// TwinCAT 3 PLC project CMoLib
// ProgramVersion: 3.1.4024.0
// libraries:
//   Tc2_Standard, * (Beckhoff Automation GmbH)
//   Tc2_System, * (Beckhoff Automation GmbH)
//   Tc2_Utilities, * (Beckhoff Automation GmbH)
//   Tc3_Module, * (Beckhoff Automation GmbH)
// project tree:
//   DUTs/ CMoDateTime.TcDUT, CMoDateTimeString.TcDUT, CMoFramework.TcDUT, CMoHalDigitalInput.TcDUT, CMoHalDigitalOutput.TcDUT, CMoInterlock.TcDUT
//   GVLs/ GVL.TcGVL
//   / PlcTask.TcTTO
//   POUs/ CMoDateTimeToString.TcPOU, CMoDiffTime.TcPOU, CMoDigitalInput.TcPOU, CMoDigitalOutput.TcPOU, CMoElapsedTime.TcPOU, CMoEvalInterlock.TcPOU, CMoGetLocalDateTime.TcPOU, CMoGetUTCDateTime.TcPOU, CMoMainRuntime.TcPOU, CMoRandom.TcPOU, MAIN.TcPOU
// real-time tasks:
//   TASK PlcTask: cycle T#5ms, priority 20, ADS port 350

CONFIGURATION CMoLib
    RESOURCE PLC ON TwinCAT3
        TASK PlcTask(INTERVAL := T#5ms, PRIORITY := 20);
        PROGRAM MAIN WITH PlcTask : MAIN;
    END_RESOURCE
END_CONFIGURATION

// ---- DUTs/CMoDateTime.TcDUT
// CMoDateTime — Date and Time Structure
// CMo Library v1.0 — Cristian Mori
// TwinCAT / IEC 61131-3 Structured Text

TYPE CMoDateTime :
STRUCT
    RawDateTime     : ARRAY[0..6] OF DINT;  // Platform-native wall clock data
    Year            : DINT;
    Month           : DINT;     // 1-12
    Day             : DINT;     // 1-31
    Hour            : DINT;     // 0-23
    Minute          : DINT;     // 0-59
    Second          : DINT;     // 0-59
    MicroSecond     : DINT;     // 0-999999
    IsLocal         : BOOL;     // TRUE = local time, FALSE = UTC
END_STRUCT
END_TYPE

// ---- DUTs/CMoDateTimeString.TcDUT
// CMoDateTimeString — HMI-Readable Date/Time Strings
// CMo Library v1.0 — Cristian Mori

TYPE CMoDateTimeString :
STRUCT
    TimeString      : STRING(16);   // "HH:MM:SS"
    DateString      : STRING(16);   // "YYYY-MM-DD"
    HMIString       : STRING(32);   // "YYYY-MM-DD HH:MM:SS"
END_STRUCT
END_TYPE

// ---- DUTs/CMoFramework.TcDUT
// CMoCommon — Shared System Context
// CMo Library v1.0 — Cristian Mori
//
// One instance per PLC. Passed as VAR_IN_OUT to every FB.
// Temp* fields are scratch accumulators: reset each scan by CMoMasterTask,
// set by individual FBs, then latched into final fields next scan.

TYPE CMoFramework :
STRUCT
    // ---- Alarm rollup flags ----
    AnyAudibleOn            : BOOL;
    AnyAudibleOnLastScan        : BOOL;
    AnyAlarmActive          : BOOL;
    AnyAlarmActiveLastScan      : BOOL;
    AnyWarningActive        : BOOL;
    AnyWarningActiveLastScan    : BOOL;
    AnyFaultActive          : BOOL;
    AnyFaultActiveLastScan      : BOOL;
    AnyCriticalActive       : BOOL;
    AnyCriticalActiveLastScan   : BOOL;

    // ---- Simulation / Hand detection ----
    AnySimulationOn         : BOOL;
    AnySimulationOnLastScan     : BOOL;
    AnyHandOn               : BOOL;
    AnyHandOnLastScan           : BOOL;

    // ---- HMI commands ----
    SilenceCmd              : BOOL;     // HMI silence button (momentary)
    GlobalAlmRstCmd         : BOOL;     // HMI global alarm reset (momentary)
    GlobalAlmRstEn          : BOOL;     // Enable global alarm reset

    // ---- System modes ----
    SimulationEnabled       : BOOL;     // Master simulation enable
    EmulationEnabled        : BOOL;     // Running on emulated controller
    MaintenanceEnabled      : BOOL;     // Enables Hand mode

    // ---- Tick timers (pulse TRUE for one scan) ----
    Tick100ms               : BOOL;
    Tick1s                  : BOOL;
    Tick10s                 : BOOL;

    // ---- Blinker signals (toggle on/off) ----
	Blink100ms				: BOOL;
    Blink250ms              : BOOL;
    Blink500ms              : BOOL;
    Blink1s                 : BOOL;
    Blink2s                 : BOOL;

    // ---- System flags ----
    InhibitAlarms           : BOOL;     // Corporate alarm inhibit
    AlwaysTrue              : BOOL;     // Constant TRUE
    AlwaysFalse             : BOOL;     // Constant FALSE
  

    // ---- Counters ----
    ApplicationCount        : DINT;
    AlarmCount              : INT;
    TempAlarmCount          : INT;
    FreeRunningTimer        : DINT;     // Free-running ms counter
    LastRandomSeed          : DINT;
	Random 					: REAL;
    CycleTime               : REAL;     // Last scan time (seconds)

    // ---- Group-level alarm rollups (512 groups as bit arrays) ----
    InhibitAlarmGroups              : ARRAY[0..15] OF DWORD;

    // ---- Date/Time ----
    CurrentUTCDateTime      : CMoDateTime;
    CurrentLocalDateTime    : CMoDateTime;
    CurrentUTCString        : CMoDateTimeString;
    CurrentLocalString      : CMoDateTimeString;

    // ---- Spare HAL instances ----
    NotUsedDI                 : CMoHALDigitalInput;
    NotUsedDO                 : CMoHALDigitalOutput;

    // ---- Module status config ----
    ModuleStatusMinInterval         : DINT := 5000;     // ms between checks
    ModuleStatusRandomDistribution  : DINT := 2000;     // ms random spread
    ModuleStatusGraceTime           : DINT := 30000;    // ms before declaring lost
END_STRUCT
END_TYPE

// ---- DUTs/CMoHalDigitalInput.TcDUT
// CMoHALDigitalInput — Digital Input Hardware Abstraction Layer
// CMo Library v1.0 — Cristian Mori
//
// THE CORE RULE: Business logic reads .Value only.
//
// Three signal modes:
//   Normal:     Value follows hardware Input (optionally inverted, debounced)
//   Simulation: Value follows SimInput (per-signal, for brownfield testing)
//   Hand:       Value follows HandValue (operator override from HMI)

TYPE CMoHALDigitalInput :
STRUCT
    // --- Raw hardware ---
    Input               : BOOL;     // Raw hardware input (written by device driver)
    QualityInput        : BOOL;     // Hardware health from module status (TRUE = good)

    // --- Simulation ---
    SimInput            : BOOL;     // Simulation input (written by twin/test)
    EnableSimulation    : BOOL;     // Enable simulation for this point
    SimulationIsActive  : BOOL;     // Computed: EnableSimulation AND Common.SimulationEnabled

    // --- Hand (manual override) ---
    HandValue           : BOOL;     // Manual override value (set from HMI)
    EnableHand          : BOOL;     // Enable hand mode for this point
    HandIsActive        : BOOL;     // Computed: EnableHand AND Common.MaintenanceEnabled

    // --- THE OUTPUT ---
    Value               : BOOL;     // Conditioned, filtered, mode-selected result

    // --- Configuration ---
    Inverted            : BOOL;     // Invert input polarity
    BadQualityValue     : BOOL;     // Value to use when quality is bad (safe state)
    EnableDelay         : BOOL;     // Enable debounce filtering
    IsSpare             : BOOL;     // Mark as spare (bypasses quality, forces sim)
    InFilterOnTimeMsec  : DINT;     // On-delay debounce (milliseconds)
    InFilterOffTimeMsec : DINT;     // Off-delay debounce (milliseconds)

    // --- Computed status ---
    PointQuality        : BOOL;     // Computed quality (good if hw OK or sim active)
    RisingEdge          : BOOL;     // One-shot pulse on Value 0 to 1
    FallingEdge         : BOOL;     // One-shot pulse on Value 1 to 0

    // --- Self-documenting ---
    Name                : STRING(28);
END_STRUCT
END_TYPE

// ---- DUTs/CMoHalDigitalOutput.TcDUT
// CMoHALDigitalOutput — Digital Output Hardware Abstraction Layer
// CMo Library v1.0 — Cristian Mori
//
// Business logic writes .Value. The FB handles inversion, hand mode,
// simulation capture, and quality gating before driving physical output.

TYPE CMoHALDigitalOutput :
STRUCT
    // --- Physical output ---
    Output              : BOOL;     // Physical output (written by FB to hardware)
    QualityInput        : BOOL;     // Hardware health (TRUE = good)

    // --- Simulation ---
    SimOutput           : BOOL;     // Shadow output for twin consumption during sim
    EnableSimulation    : BOOL;     // Enable simulation for this point
    SimulationIsActive  : BOOL;     // Computed: EnableSimulation AND Common.SimulationEnabled

    // --- Hand (manual override) ---
    HandValue           : BOOL;     // Manual override value (set from HMI)
    EnableHand          : BOOL;     // Enable hand mode for this point
    HandIsActive        : BOOL;     // Computed: EnableHand AND Common.MaintenanceEnabled

    // --- THE INPUT (business logic writes this) ---
    Value               : BOOL;     // Business logic command

    // --- Configuration ---
    Inverted            : BOOL;     // Invert output polarity
    BadQualityValue     : BOOL;     // Value when quality is bad (safe state)
    IsSpare             : BOOL;     // Mark as spare

    // --- Computed status ---
    PointQuality        : BOOL;     // Computed quality

    // --- Self-documenting ---
    Name                : STRING(28);
END_STRUCT
END_TYPE

// ---- DUTs/CMoInterlock.TcDUT
// CMoInterlock — Interlock Condition Structure
// CMo Library v1.0 — Cristian Mori
//
// Up to 16 AND conditions. All must be TRUE for interlock to pass.
// FirstOut: which condition dropped first (root cause).
// Per-condition bypass from HMI with bypass alarm.

TYPE CMoInterlock :
STRUCT
    // Configuration
    PointCount          : INT := 4;     // Number of active conditions (1-16)

    // Condition inputs (set by business logic each scan)
    Condition           : ARRAY[0..15] OF BOOL;

    // Per-condition bypass (set from HMI)
    Bypass              : ARRAY[0..15] OF BOOL;

    // Outputs
    OK                  : BOOL;     // All active conditions met (or bypassed)
    InBypass            : BOOL;     // At least one condition is bypassed
    BypassAlarm         : BOOL;     // Alarm: operating with bypassed conditions

    // First-out tracking
    FirstOut            : INT := -1; // Index of first condition to drop (-1 = none)

    // Per-condition status (for HMI popup)
    ConditionMet        : ARRAY[0..15] OF BOOL;  // Condition OR its bypass
    ConditionFaulted    : ARRAY[0..15] OF BOOL;  // Failed AND not bypassed

    // Self-documenting names
    Name                : STRING(28);
    ConditionName       : ARRAY[0..15] OF STRING(28);
END_STRUCT
END_TYPE

// ---- GVLs/GVL.TcGVL
{attribute 'qualified_only'}
VAR_GLOBAL
    Framework       : CMoFramework;
	
	DI_PartPresent  : CMoHALDigitalInput;
    DI_GuardClosed  : CMoHALDigitalInput;
    DO_MotorRun     : CMoHALDigitalOutput;
    Interlock_Motor : CMoInterlock;
END_VAR

// ---- POUs/MAIN.TcPOU
PROGRAM MAIN
VAR
	fbMainRuntime    : CMoMainRuntime;
	fbInterlock 	 : CMoEvalInterlock;
	fbPartPresent	 : CMoDigitalInput;
	fbGuardClosed	 : CMoDigitalInput;
	fbMotorRun		 : CMoDigitalOutput;
	fDiffTime	     : CMoDiffTime;
	SimPartPresent	 : BOOL;
	SimGuardClosed	 : BOOL;
	saveStart: BOOL;
	StartDate: CMoDateTime;
	saveEnd: BOOL;
	EndDate: CMoDateTime;
	totSec: DINT;
	TotuSec: DINT;
END_VAR

// Heartbeat: always first
fbMainRuntime(Framework := GVL.Framework);

// Enable simulation globally
GVL.Framework.SimulationEnabled := TRUE;

GVL.Framework.SimulationEnabled := TRUE;

// --- Part Present sensor ---
GVL.DI_PartPresent.EnableSimulation := TRUE;
GVL.DI_PartPresent.SimInput := SimPartPresent;
GVL.DI_PartPresent.Name := 'Part Present';

fbPartPresent(
    HAL := GVL.DI_PartPresent,
    DeviceInput := FALSE,
    QualityInput := TRUE,
    Framework := GVL.Framework
);

// --- Guard Door sensor ---
GVL.DI_GuardClosed.EnableSimulation := TRUE;
GVL.DI_GuardClosed.SimInput := SimGuardClosed;
GVL.DI_GuardClosed.Name := 'Guard Closed';

fbGuardClosed(
    HAL := GVL.DI_GuardClosed,
    DeviceInput := FALSE,
    QualityInput := TRUE,
    Framework := GVL.Framework
);

// --- Interlock ---
GVL.Interlock_Motor.PointCount := 2;
GVL.Interlock_Motor.ConditionName[0] := 'Part Present';
GVL.Interlock_Motor.ConditionName[1] := 'Guard Closed';
GVL.Interlock_Motor.Condition[0] := GVL.DI_PartPresent.Value;
GVL.Interlock_Motor.Condition[1] := GVL.DI_GuardClosed.Value;

fbInterlock(Ilk := GVL.Interlock_Motor);

// --- Business logic: .Value only ---
GVL.DO_MotorRun.EnableSimulation := TRUE;
GVL.DO_MotorRun.Value := GVL.Interlock_Motor.OK;
GVL.DO_MotorRun.Name := 'Motor Run';

fbMotorRun(
    HAL := GVL.DO_MotorRun,
    QualityInput := TRUE,
    Framework := GVL.Framework
);

IF saveStart THEN
	StartDate :=  GVL.Framework.CurrentUTCDateTime;
END_IF

IF saveEnd THEN
	EndDate :=  GVL.Framework.CurrentUTCDateTime;
END_IF

fDiffTime(StartTime := StartDate,EndTime := EndDate);
totSec:=fDiffTime.TotalSeconds;
totuSec:=fDiffTime.TotalMicroseconds;

END_PROGRAM

// ---- POUs/CMoMainRuntime.TcPOU
FUNCTION_BLOCK CMoMainRuntime
VAR_INPUT
END_VAR
VAR_OUTPUT
END_VAR
VAR_IN_OUT
    Framework       : CMoFramework;
END_VAR
VAR
    // Tick timers
    tmTick100ms     : TON;
    tmTick1s        : TON;
    tmTick10s       : TON;

    // Blinker timers
    tmBlink100ms    : TON;
    tmBlink250ms    : TON;
    tmBlink500ms    : TON;
    tmBlink1s       : TON;
    tmBlink2s       : TON;
    bState100ms     : BOOL;
    bState250ms     : BOOL;
    bState500ms     : BOOL;
    bState1s        : BOOL;
    bState2s        : BOOL;

    // DateTime FBs
    fbGetLocal      : CMoGetLocalDateTime;
    fbGetUTC        : CMoGetUTCDateTime;
    fbLocalToStr    : CMoDateTimeToString;
    fbUTCToStr      : CMoDateTimeToString;
	
	    // Scan time measurement
    fbScanTime      : CMoElapsedTime;
    bScanRunning    : BOOL;
 
    // Random number generator
    fbRandom        : CMoRandom;
END_VAR

// =============================================================================
// CMoMainRuntime — System Heartbeat
// CMo Library v1.0
// =============================================================================
// Call ONCE per scan, FIRST in the task. Responsible for:
//   - Measuring scan cycle time (via CMoElapsedTime)
//   - Generating tick timers (100ms, 1s, 10s)
//   - Generating blinker signals (100ms, 250ms, 500ms, 1s, 2s)
//   - Latching LastScan accumulators into final alarm/sim/hand rollups
//   - Resetting LastScan accumulators for the new scan
//   - Generating random number (via CMoRandom)
//   - Updating local and UTC date/time with formatted strings
//   - Setting constants (AlwaysTrue, AlwaysFalse)
//   - Incrementing free-running timer
//
// The LastScan pattern:
//   MainRuntime resets all *LastScan fields at start of scan.
//   Individual CMoAlarm/CMoDigitalInput FBs SET them during the scan.
//   MainRuntime copies LastScan -> final at the NEXT call.
//   This eliminates execution order dependencies.
//
// Usage:
//   fbRuntime(Framework := GVL.Framework);  // first line of MAIN
// =============================================================================

// =================================================================
// Scan time measurement: stop previous, read result, start new
// =================================================================
IF bScanRunning THEN
    // Stop the timer from last scan
    fbScanTime(Start := FALSE, Stop := TRUE, Reset := FALSE);
    Framework.CycleTime := fbScanTime.ElapsedMs;
    // Reset and start fresh for this scan
    fbScanTime(Start := FALSE, Stop := FALSE, Reset := TRUE);
    fbScanTime(Start := TRUE, Stop := FALSE, Reset := FALSE);
ELSE
    // First scan: just start
    fbScanTime(Start := TRUE, Stop := FALSE, Reset := FALSE);
    bScanRunning := TRUE;
END_IF;

// =================================================================
// Latch previous scan accumulators into final outputs
// =================================================================
Framework.AnyAudibleOn       := Framework.AnyAudibleOnLastScan;
Framework.AnyAlarmActive     := Framework.AnyAlarmActiveLastScan;
Framework.AnyWarningActive   := Framework.AnyWarningActiveLastScan;
Framework.AnyFaultActive     := Framework.AnyFaultActiveLastScan;
Framework.AnyCriticalActive  := Framework.AnyCriticalActiveLastScan;
Framework.AnySimulationOn    := Framework.AnySimulationOnLastScan;
Framework.AnyHandOn          := Framework.AnyHandOnLastScan;
Framework.AlarmCount         := Framework.TempAlarmCount;

// =================================================================
// Reset scratch for this scan
// =================================================================
Framework.AnyAudibleOnLastScan      := FALSE;
Framework.AnyAlarmActiveLastScan    := FALSE;
Framework.AnyWarningActiveLastScan  := FALSE;
Framework.AnyFaultActiveLastScan    := FALSE;
Framework.AnyCriticalActiveLastScan := FALSE;
Framework.AnySimulationOnLastScan   := FALSE;
Framework.AnyHandOnLastScan         := FALSE;
Framework.TempAlarmCount            := 0;

// =================================================================
// Constants
// =================================================================
Framework.AlwaysTrue  := TRUE;
Framework.AlwaysFalse := FALSE;

// =================================================================
// Random number generator
// =================================================================
fbRandom(Seed := Framework.LastRandomSeed);
Framework.Random := fbRandom.Out;
Framework.LastRandomSeed := fbRandom.NewSeed;

// =================================================================
// Ticks: pulse TRUE for one scan at each interval
// =================================================================
tmTick100ms(IN := TRUE, PT := T#100MS);
Framework.Tick100ms := tmTick100ms.Q;
IF tmTick100ms.Q THEN
    tmTick100ms(IN := FALSE, PT := T#100MS);
END_IF;

tmTick1s(IN := TRUE, PT := T#1S);
Framework.Tick1s := tmTick1s.Q;
IF tmTick1s.Q THEN
    tmTick1s(IN := FALSE, PT := T#1S);
END_IF;

tmTick10s(IN := TRUE, PT := T#10S);
Framework.Tick10s := tmTick10s.Q;
IF tmTick10s.Q THEN
    tmTick10s(IN := FALSE, PT := T#10S);
END_IF;

// =================================================================
// Blinkers: toggle state at each interval
// =================================================================
tmBlink100ms(IN := TRUE, PT := T#100MS);
IF tmBlink100ms.Q THEN
    bState100ms := NOT bState100ms;
    tmBlink100ms(IN := FALSE, PT := T#100MS);
END_IF;
Framework.Blink100ms := bState100ms;

tmBlink250ms(IN := TRUE, PT := T#250MS);
IF tmBlink250ms.Q THEN
    bState250ms := NOT bState250ms;
    tmBlink250ms(IN := FALSE, PT := T#250MS);
END_IF;
Framework.Blink250ms := bState250ms;

tmBlink500ms(IN := TRUE, PT := T#500MS);
IF tmBlink500ms.Q THEN
    bState500ms := NOT bState500ms;
    tmBlink500ms(IN := FALSE, PT := T#500MS);
END_IF;
Framework.Blink500ms := bState500ms;

tmBlink1s(IN := TRUE, PT := T#1S);
IF tmBlink1s.Q THEN
    bState1s := NOT bState1s;
    tmBlink1s(IN := FALSE, PT := T#1S);
END_IF;
Framework.Blink1s := bState1s;

tmBlink2s(IN := TRUE, PT := T#2S);
IF tmBlink2s.Q THEN
    bState2s := NOT bState2s;
    tmBlink2s(IN := FALSE, PT := T#2S);
END_IF;
Framework.Blink2s := bState2s;

// =================================================================
// Free-running timer
// =================================================================
Framework.FreeRunningTimer := Framework.FreeRunningTimer + 1;

// =================================================================
// Date/Time: read local and UTC, format strings
// =================================================================
fbGetLocal(DateTime := Framework.CurrentLocalDateTime);
fbGetUTC(DateTime := Framework.CurrentUTCDateTime);

fbLocalToStr(
    DateTime := Framework.CurrentLocalDateTime,
    DateTimeString := Framework.CurrentLocalString
);
fbUTCToStr(
    DateTime := Framework.CurrentUTCDateTime,
    DateTimeString := Framework.CurrentUTCString
);

END_FUNCTION_BLOCK

// ---- POUs/CMoGetLocalDateTime.TcPOU
FUNCTION_BLOCK CMoGetLocalDateTime
VAR_INPUT
END_VAR
VAR_OUTPUT
END_VAR
VAR_IN_OUT
    DateTime        : CMoDateTime;
END_VAR
VAR
	fbLocalTime     : FB_LocalSystemTime := (bEnable := TRUE, dwCycle := 1);
END_VAR

// =============================================================================
// CMoGetLocalDateTime — Read Local System Time (Beckhoff)
// CMo Library v1.0
// Requires: Tc2_Utilities library
// =============================================================================
// Reads the local Windows system time via FB_LocalSystemTime and
// maps TIMESTRUCT fields into CMoDateTime.
//
// Must be called cyclically. Called internally by CMoMainRuntime
// every scan.
//
// Usage:
//   fbLocal(DateTime := Framework.CurrentLocalDateTime);
// =============================================================================

fbLocalTime();
IF fbLocalTime.bValid THEN
    DateTime.Year        := WORD_TO_DINT(fbLocalTime.systemTime.wYear);
    DateTime.Month       := WORD_TO_DINT(fbLocalTime.systemTime.wMonth);
    DateTime.Day         := WORD_TO_DINT(fbLocalTime.systemTime.wDay);
    DateTime.Hour        := WORD_TO_DINT(fbLocalTime.systemTime.wHour);
    DateTime.Minute      := WORD_TO_DINT(fbLocalTime.systemTime.wMinute);
    DateTime.Second      := WORD_TO_DINT(fbLocalTime.systemTime.wSecond);
    DateTime.MicroSecond := WORD_TO_DINT(fbLocalTime.systemTime.wMilliseconds) * 1000;
    DateTime.IsLocal     := TRUE;
END_IF;

END_FUNCTION_BLOCK

// ---- POUs/CMoGetUTCDateTime.TcPOU
FUNCTION_BLOCK CMoGetUTCDateTime
VAR_IN_OUT
    DateTime        : CMoDateTime;
END_VAR
VAR_INPUT
END_VAR
VAR_OUTPUT
END_VAR
VAR
	fbLocalTime     : FB_LocalSystemTime := (bEnable := TRUE, dwCycle := 1);
    fbToUTC         : FB_TzSpecificLocalTimeToSystemTime;
    fbGetTZ         : FB_GetTimeZoneInformation;
    tzInfo          : ST_TimeZoneInformation;
    utcTime         : TIMESTRUCT;
    bTzValid        : BOOL;
END_VAR

// =============================================================================
// CMoGetUTCDateTime — Read UTC System Time (Beckhoff)
// CMo Library v1.0
// Requires: Tc2_Utilities library
// =============================================================================
// Reads the local Windows system time via FB_LocalSystemTime, then
// converts to UTC using FB_TzSpecificLocalTimeToSystemTime with
// timezone info from FB_GetTimeZoneInformation.
//
// Must be called cyclically. Populates a CMoDateTime with UTC fields.
// Called internally by CMoMainRuntime every scan.
//
// Usage:
//   fbUTC(DateTime := Framework.CurrentUTCDateTime);
// =============================================================================

// Get local time (must call cyclically)
fbLocalTime();

// Get timezone info (for local-to-UTC conversion)
fbGetTZ(
    sNetID := '',
    bExecute := NOT bTzValid,
    tTimeout := DEFAULT_ADS_TIMEOUT
);
IF NOT fbGetTZ.bBusy AND NOT fbGetTZ.bError THEN
    tzInfo := fbGetTZ.tzInfo;
    bTzValid := TRUE;
END_IF;

// Convert local to UTC
IF fbLocalTime.bValid AND bTzValid THEN
    fbToUTC(
        in := fbLocalTime.systemTime,
        tzInfo := tzInfo
    );
    utcTime := fbToUTC.out;

    DateTime.Year        := WORD_TO_DINT(utcTime.wYear);
    DateTime.Month       := WORD_TO_DINT(utcTime.wMonth);
    DateTime.Day         := WORD_TO_DINT(utcTime.wDay);
    DateTime.Hour        := WORD_TO_DINT(utcTime.wHour);
    DateTime.Minute      := WORD_TO_DINT(utcTime.wMinute);
    DateTime.Second      := WORD_TO_DINT(utcTime.wSecond);
    DateTime.MicroSecond := WORD_TO_DINT(utcTime.wMilliseconds) * 1000;
    DateTime.IsLocal     := FALSE;
END_IF;

END_FUNCTION_BLOCK

// ---- POUs/CMoDateTimeToString.TcPOU
FUNCTION_BLOCK CMoDateTimeToString
VAR_INPUT
    DateTime        : CMoDateTime;
END_VAR
VAR_IN_OUT
    DateTimeString  : CMoDateTimeString;
END_VAR
VAR_OUTPUT
END_VAR
VAR
	sYear           : STRING(4);
    sMonth          : STRING(2);
    sDay            : STRING(2);
    sHour           : STRING(2);
    sMinute         : STRING(2);
    sSecond         : STRING(2);
END_VAR

// =============================================================================
// CMoDateTimeToString — Format DateTime for HMI Display
// CMo Library v1.0
// =============================================================================
// Converts CMoDateTime fields into zero-padded human-readable strings:
//   TimeString: "HH:MM:SS"
//   DateString: "YYYY-MM-DD"
//   HMIString:  "YYYY-MM-DD HH:MM:SS"
//
// Usage:
//   fbFmt(DateTime := myTime, DateTimeString := myStrings);
//   // myStrings.HMIString now holds "2026-04-09 14:30:05"
// =============================================================================

sYear := DINT_TO_STRING(DateTime.Year);

IF DateTime.Month < 10 THEN
    sMonth := CONCAT('0', DINT_TO_STRING(DateTime.Month));
ELSE
    sMonth := DINT_TO_STRING(DateTime.Month);
END_IF;

IF DateTime.Day < 10 THEN
    sDay := CONCAT('0', DINT_TO_STRING(DateTime.Day));
ELSE
    sDay := DINT_TO_STRING(DateTime.Day);
END_IF;

IF DateTime.Hour < 10 THEN
    sHour := CONCAT('0', DINT_TO_STRING(DateTime.Hour));
ELSE
    sHour := DINT_TO_STRING(DateTime.Hour);
END_IF;

IF DateTime.Minute < 10 THEN
    sMinute := CONCAT('0', DINT_TO_STRING(DateTime.Minute));
ELSE
    sMinute := DINT_TO_STRING(DateTime.Minute);
END_IF;

IF DateTime.Second < 10 THEN
    sSecond := CONCAT('0', DINT_TO_STRING(DateTime.Second));
ELSE
    sSecond := DINT_TO_STRING(DateTime.Second);
END_IF;

DateTimeString.TimeString := CONCAT(CONCAT(CONCAT(CONCAT(sHour, ':'), sMinute), ':'), sSecond);
DateTimeString.DateString := CONCAT(CONCAT(CONCAT(CONCAT(sYear, '-'), sMonth), '-'), sDay);
DateTimeString.HMIString  := CONCAT(CONCAT(DateTimeString.DateString, ' '), DateTimeString.TimeString);

END_FUNCTION_BLOCK

// ---- POUs/CMoElapsedTime.TcPOU
FUNCTION_BLOCK CMoElapsedTime
VAR_INPUT
    Start           : BOOL;         // Begin measurement (rising edge)
    Stop            : BOOL;         // End measurement (rising edge)
    Reset           : BOOL;         // Clear measurement
END_VAR
VAR_OUTPUT
    ElapsedMs       : REAL;         // Result in milliseconds
    Running         : BOOL;         // TRUE while measuring
END_VAR
VAR
    PrevStart       : BOOL;         // Edge detection for Start
    PrevStop        : BOOL;         // Edge detection for Stop
    tmRun           : TON;          // Internal timer
    Capturing       : BOOL;         // Measurement in progress
END_VAR

// =============================================================================
// CMoElapsedTime — Elapsed Time Measurement
// CMo Library v1.0
// =============================================================================
// Measures elapsed time between Start and Stop rising edges.
// Uses a TON timer internally for millisecond-resolution measurement.
// Live readout available via ElapsedMs while Running is TRUE.
//
// Usage:
//   myTimer(Start := TRUE);       // Begin measurement
//   // ... code or scans pass ...
//   myTimer(Stop := TRUE);        // End measurement
//   result := myTimer.ElapsedMs;  // Read duration in ms
//   myTimer(Reset := TRUE);       // Clear for next use
// =============================================================================

// =================================================================
// Reset: clear everything
// =================================================================
IF Reset THEN
    ElapsedMs := 0.0;
    Running := FALSE;
    Capturing := FALSE;
    RETURN;
END_IF;

// =================================================================
// Start on rising edge: reset timer and begin capturing
// =================================================================
IF Start AND NOT PrevStart THEN
    Capturing := TRUE;
    Running := TRUE;
    tmRun(IN := FALSE, PT := T#49D);   // Reset timer (49 day max range)
END_IF;
PrevStart := Start;

// =================================================================
// Accumulate while running: keep timer alive, update live readout
// =================================================================
IF Capturing THEN
    tmRun(IN := TRUE, PT := T#49D);
    ElapsedMs := TIME_TO_REAL(tmRun.ET);
END_IF;

// =================================================================
// Stop on rising edge: freeze result
// =================================================================
IF Stop AND NOT PrevStop AND Capturing THEN
    ElapsedMs := TIME_TO_REAL(tmRun.ET);
    Capturing := FALSE;
    Running := FALSE;
END_IF;
PrevStop := Stop;

END_FUNCTION_BLOCK

// ---- POUs/CMoRandom.TcPOU
FUNCTION_BLOCK CMoRandom
VAR_INPUT
    Seed            : DINT := 48271;
END_VAR
VAR_OUTPUT
    Out             : REAL;
    NewSeed         : DINT;
END_VAR

// =============================================================================
// CMoRandom — Random Number Generator
// CMo Library v1.0
// =============================================================================
// Park-Miller linear congruential generator.
// Outputs a REAL between 0.0 and 1.0.
//
// Feed Seed from Framework.LastRandomSeed, write NewSeed back after call.
// Called internally by CMoMainRuntime every scan.
//
// Usage:
//   fbRandom(Seed := Framework.LastRandomSeed);
//   Framework.Random := fbRandom.Out;
//   Framework.LastRandomSeed := fbRandom.NewSeed;
// =============================================================================

// Ensure positive seed
IF Seed <= 0 THEN
    Seed := 1;
END_IF;
 
// Park-Miller LCG: next = (seed * 16807) MOD 2147483647
// Classic "Minimal Standard" PRNG, different algorithm from typical PLC implementations
NewSeed := (Seed MOD 127773) * 16807 - (Seed / 127773) * 2836;
IF NewSeed <= 0 THEN
    NewSeed := NewSeed + 2147483647;
END_IF;
 
Out := DINT_TO_REAL(NewSeed) / 2147483647.0;

END_FUNCTION_BLOCK

// ---- POUs/CMoEvalInterlock.TcPOU
FUNCTION_BLOCK CMoEvalInterlock
VAR_IN_OUT
    Ilk             : CMoInterlock;
END_VAR
VAR
    i               : INT;
    AllMet          : BOOL;
    AnyBypassed     : BOOL;
    FirstDropped    : INT;
    PrevOK          : BOOL;
END_VAR

// =================================================================
// Clamp PointCount
// =================================================================
IF Ilk.PointCount < 1 THEN
    Ilk.PointCount := 1;
ELSIF Ilk.PointCount > 16 THEN
    Ilk.PointCount := 16;
END_IF;

// =================================================================
// Evaluate each condition
// =================================================================
AllMet := TRUE;
AnyBypassed := FALSE;
FirstDropped := -1;

FOR i := 0 TO Ilk.PointCount - 1 DO
    Ilk.ConditionMet[i] := Ilk.Condition[i] OR Ilk.Bypass[i];
    Ilk.ConditionFaulted[i] := NOT Ilk.Condition[i] AND NOT Ilk.Bypass[i];

    IF Ilk.Bypass[i] THEN
        AnyBypassed := TRUE;
    END_IF;

    IF Ilk.ConditionFaulted[i] AND FirstDropped = -1 THEN
        FirstDropped := i;
    END_IF;

    IF NOT Ilk.ConditionMet[i] THEN
        AllMet := FALSE;
    END_IF;
END_FOR;

// Clear unused conditions
FOR i := Ilk.PointCount TO 15 DO
    Ilk.ConditionMet[i] := TRUE;
    Ilk.ConditionFaulted[i] := FALSE;
END_FOR;

// =================================================================
// Outputs
// =================================================================
PrevOK := Ilk.OK;
Ilk.OK := AllMet;
Ilk.InBypass := AnyBypassed;
Ilk.BypassAlarm := AnyBypassed;

// =================================================================
// FirstOut: latch on OK->NOT OK transition
// =================================================================
IF NOT Ilk.OK AND PrevOK THEN
    Ilk.FirstOut := FirstDropped;
ELSIF Ilk.OK THEN
    Ilk.FirstOut := -1;
END_IF;

END_FUNCTION_BLOCK

// ---- POUs/CMoDigitalInput.TcPOU
FUNCTION_BLOCK CMoDigitalInput
VAR_IN_OUT
    HAL             : CMoHALDigitalInput;
    Framework       : CMoFramework;
END_VAR
VAR_INPUT
    DeviceInput     : BOOL;
    QualityInput    : BOOL;
END_VAR
VAR
    ConditionedInput    : BOOL;
    DebouncedValue      : BOOL;
    OnDelayTimer        : TON;
    OffDelayTimer       : TOF;
    PrevValue           : BOOL;
    FirstScan           : BOOL := TRUE;
    ReSync              : BOOL;
    NoFilterNeeded      : BOOL;
END_VAR

// =============================================================================
// CMoDigitalInput — Digital Input Signal Conditioning
// CMo Library v1.0
// =============================================================================
// Takes a raw hardware input and produces a conditioned .Value through:
//   1. Mode determination (Normal / Simulation / Hand)
//   2. Quality evaluation (hardware health, sim, spare)
//   3. Mode selection + polarity inversion
//   4. Debounce filtering (configurable on/off delay with resync)
//   5. Hand value bumpless transfer
//   6. Quality gating (bad quality -> configurable fallback)
//   7. Edge detection (RisingEdge / FallingEdge one-shot pulses)
//
// Business logic reads .Value only. Never touch .Input, .SimInput,
// .HandValue, or any plumbing directly.
//
// Usage:
//   fbInput(
//       HAL := GVL.MyInput,
//       DeviceInput := Module1:I.Data[0],
//       QualityInput := Module1_Status.Running,
//       Framework := GVL.Framework
//   );
// =============================================================================

// =================================================================
// Mode determination
// =================================================================
HAL.HandIsActive := HAL.EnableHand AND Framework.MaintenanceEnabled;
IF HAL.HandIsActive THEN
    Framework.AnyHandOnLastScan := TRUE;
END_IF;

HAL.SimulationIsActive := HAL.EnableSimulation AND Framework.SimulationEnabled;
IF HAL.SimulationIsActive THEN
    Framework.AnySimulationOnLastScan := TRUE;
END_IF;

// =================================================================
// Point quality
// =================================================================
IF HAL.IsSpare THEN
    HAL.PointQuality := TRUE;
ELSIF HAL.SimulationIsActive THEN
    HAL.PointQuality := TRUE;
ELSE
    HAL.QualityInput := QualityInput;
    HAL.PointQuality := QualityInput;
END_IF;

// =================================================================
// Latch raw input
// =================================================================
HAL.Input := DeviceInput;

// =================================================================
// Mode selection + inversion
// =================================================================
IF HAL.SimulationIsActive THEN
    IF HAL.Inverted THEN
        ConditionedInput := NOT HAL.SimInput;
    ELSE
        ConditionedInput := HAL.SimInput;
    END_IF;
ELSE
    IF HAL.Inverted THEN
        ConditionedInput := NOT HAL.Input;
    ELSE
        ConditionedInput := HAL.Input;
    END_IF;
END_IF;

// =================================================================
// Debounce filter
// =================================================================
IF NOT HAL.EnableDelay THEN
    DebouncedValue := ConditionedInput;
    ReSync := TRUE;
ELSE
    IF HAL.InFilterOnTimeMsec < 0 THEN
        HAL.InFilterOnTimeMsec := 0;
    END_IF;
    IF HAL.InFilterOffTimeMsec < 0 THEN
        HAL.InFilterOffTimeMsec := 0;
    END_IF;

    OnDelayTimer(
        IN := ConditionedInput OR (OffDelayTimer.Q AND OnDelayTimer.Q),
        PT := DINT_TO_TIME(HAL.InFilterOnTimeMsec)
    );

    OffDelayTimer(
        IN := ConditionedInput,
        PT := DINT_TO_TIME(HAL.InFilterOffTimeMsec)
    );

    NoFilterNeeded := (ConditionedInput AND OnDelayTimer.Q)
                   OR (NOT ConditionedInput AND NOT OffDelayTimer.Q);

    IF ReSync THEN
        IF (DebouncedValue AND OnDelayTimer.Q) OR
           (NOT DebouncedValue AND NOT OnDelayTimer.Q) THEN
            ReSync := FALSE;
        END_IF;
    END_IF;

    IF ReSync OR HAL.IsSpare THEN
        DebouncedValue := ConditionedInput;
    ELSIF OnDelayTimer.Q THEN
        DebouncedValue := TRUE;
    ELSIF NOT OffDelayTimer.Q THEN
        DebouncedValue := FALSE;
    END_IF;
END_IF;

// =================================================================
// Hand value tracking (bumpless transfer)
// =================================================================
IF NOT HAL.HandIsActive THEN
    HAL.HandValue := HAL.Value;
END_IF;

// =================================================================
// Final value with quality gating
// =================================================================
IF HAL.PointQuality THEN
    IF HAL.HandIsActive THEN
        HAL.Value := HAL.HandValue;
    ELSE
        HAL.Value := DebouncedValue;
    END_IF;
ELSE
    HAL.Value := HAL.BadQualityValue;
END_IF;

// =================================================================
// Edge detection
// =================================================================
IF FirstScan THEN
    PrevValue := HAL.Value;
    HAL.RisingEdge := FALSE;
    HAL.FallingEdge := FALSE;
    FirstScan := FALSE;
ELSE
    HAL.RisingEdge  := HAL.Value AND NOT PrevValue;
    HAL.FallingEdge := NOT HAL.Value AND PrevValue;
    PrevValue := HAL.Value;
END_IF;

END_FUNCTION_BLOCK

// ---- POUs/CMoDigitalOutput.TcPOU
FUNCTION_BLOCK CMoDigitalOutput
VAR_IN_OUT
    HAL             : CMoHALDigitalOutput;
    Framework       : CMoFramework;
END_VAR
VAR_INPUT
    QualityInput    : BOOL;
END_VAR
VAR_OUTPUT
    DeviceOutput    : BOOL;
END_VAR
VAR
    ConditionedOutput   : BOOL;
    OutputWithHand      : BOOL;
END_VAR

// =============================================================================
// CMoDigitalOutput — Digital Output Signal Conditioning
// CMo Library v1.0
// =============================================================================
// Takes .Value written by business logic and produces a conditioned
// physical output through:
//   1. Mode determination (Normal / Simulation / Hand)
//   2. Quality evaluation (hardware health, sim, spare)
//   3. Polarity inversion
//   4. Hand value bumpless transfer
//   5. Hand mode selection
//   6. Simulation gating (suppress physical output, capture to .SimOutput)
//
// In simulation mode: DeviceOutput is suppressed. The digital twin
// reads .SimOutput to see what business logic commanded.
//
// Usage:
//   fbOutput(
//       HAL := GVL.MyOutput,
//       QualityInput := Module2_Status.Running,
//       Framework := GVL.Framework
//   );
//   Module2:O.Data[0] := fbOutput.DeviceOutput;
// =============================================================================

// =================================================================
// Mode determination
// =================================================================
HAL.HandIsActive := HAL.EnableHand AND Framework.MaintenanceEnabled AND NOT HAL.IsSpare;
IF HAL.HandIsActive THEN
    Framework.AnyHandOnLastScan := TRUE;
END_IF;

HAL.SimulationIsActive := HAL.EnableSimulation AND Framework.SimulationEnabled;
IF HAL.SimulationIsActive THEN
    Framework.AnySimulationOnLastScan := TRUE;
END_IF;

// =================================================================
// Point quality
// =================================================================
IF HAL.IsSpare THEN
    HAL.PointQuality := TRUE;
ELSIF HAL.SimulationIsActive THEN
    HAL.PointQuality := TRUE;
ELSE
    HAL.QualityInput := QualityInput;
    HAL.PointQuality := QualityInput;
END_IF;

// =================================================================
// Inversion
// =================================================================
IF NOT HAL.IsSpare THEN
    IF HAL.Inverted THEN
        ConditionedOutput := NOT HAL.Value;
    ELSE
        ConditionedOutput := HAL.Value;
    END_IF;
ELSE
    ConditionedOutput := FALSE;
END_IF;

// =================================================================
// Hand value tracking (bumpless transfer)
// =================================================================
IF NOT HAL.HandIsActive THEN
    HAL.HandValue := HAL.Value;
END_IF;

// =================================================================
// Hand mode selection
// =================================================================
IF HAL.HandIsActive THEN
    OutputWithHand := HAL.HandValue;
ELSE
    OutputWithHand := ConditionedOutput;
END_IF;

// =================================================================
// Simulation gating
// =================================================================
IF HAL.SimulationIsActive THEN
    DeviceOutput := FALSE;
ELSE
    DeviceOutput := OutputWithHand;
END_IF;

HAL.SimOutput := OutputWithHand;
HAL.Output := DeviceOutput;

END_FUNCTION_BLOCK

// ---- POUs/CMoDiffTime.TcPOU
FUNCTION_BLOCK CMoDiffTime
VAR_INPUT
    StartTime : CMoDateTime;
    EndTime   : CMoDateTime;
END_VAR
VAR_OUTPUT
    Result            : CMoDateTime;
    TotalSeconds      : DINT;
    TotalMicroseconds : DINT;
END_VAR
VAR
    jdnStart : DINT;
    jdnEnd   : DINT;
    a        : DINT;
    y        : DINT;
    m        : DINT;
    diffDays : DINT;
    diffUs   : DINT;
    diffSec  : DINT;
    diffMin  : DINT;
    diffHr   : DINT;
END_VAR

// =============================================================================
// CMoDiffTime — DateTime Subtraction via Julian Day Number
// CMo Library v1.0
// =============================================================================
// Computes (EndTime - StartTime) using Julian Day Number conversion.
// Converts both dates to JDN (integer day count), subtracts, then
// handles sub-day time remainder with borrow propagation.
//
// This is mathematically correct for all valid dates regardless of
// month lengths, leap years, or century boundaries.
//
// JDN formula (all integer math):
//   a := (14 - Month) / 12
//   y := Year + 4800 - a
//   m := Month + 12*a - 3
//   JDN := Day + (153*m + 2)/5 + 365*y + y/4 - y/100 + y/400 - 32045
//
// Usage:
//   fbDiff(StartTime := tStart, EndTime := tEnd);
//   elapsed := fbDiff.TotalSeconds;
// =============================================================================


 
// JDN for StartTime
a := (14 - StartTime.Month) / 12;
y := StartTime.Year + 4800 - a;
m := StartTime.Month + 12 * a - 3;
jdnStart := StartTime.Day + (153 * m + 2) / 5 + 365 * y + y / 4 - y / 100 + y / 400 - 32045;
 
// JDN for EndTime
a := (14 - EndTime.Month) / 12;
y := EndTime.Year + 4800 - a;
m := EndTime.Month + 12 * a - 3;
jdnEnd := EndTime.Day + (153 * m + 2) / 5 + 365 * y + y / 4 - y / 100 + y / 400 - 32045;
 
// Day difference
diffDays := jdnEnd - jdnStart;
 
// Sub-day difference with borrow propagation
diffUs := EndTime.MicroSecond - StartTime.MicroSecond;
IF diffUs < 0 THEN
    diffUs := diffUs + 1000000;
    diffSec := -1;
ELSE
    diffSec := 0;
END_IF;
 
diffSec := diffSec + EndTime.Second - StartTime.Second;
IF diffSec < 0 THEN
    diffSec := diffSec + 60;
    diffMin := -1;
ELSE
    diffMin := 0;
END_IF;
 
diffMin := diffMin + EndTime.Minute - StartTime.Minute;
IF diffMin < 0 THEN
    diffMin := diffMin + 60;
    diffHr := -1;
ELSE
    diffHr := 0;
END_IF;
 
diffHr := diffHr + EndTime.Hour - StartTime.Hour;
IF diffHr < 0 THEN
    diffHr := diffHr + 24;
    diffDays := diffDays - 1;
END_IF;
 
// Populate result
Result.Year := 0;
Result.Month := 0;
Result.Day := diffDays;
Result.Hour := diffHr;
Result.Minute := diffMin;
Result.Second := diffSec;
Result.MicroSecond := diffUs;
Result.IsLocal := FALSE;
 
// Convenience totals
TotalSeconds := diffSec + (diffMin * 60) + (diffHr * 3600) + (diffDays * 86400);
TotalMicroseconds := diffUs;

END_FUNCTION_BLOCK
